// TIA Portal V21 export
// export: Created 2026-11-10T19:11:41.578579Z, ExportSetting WithDefaults, DisplayName Totally Integrated Automation Portal, DisplayVersion V21 Update 3, DisplayName STEP 7 Professional, DisplayVersion V21 Update 3, DisplayName STEP 7 Safety, DisplayVersion V21, DisplayName Tech WebApplication, DisplayVersion V21, DisplayName WinCC Basic/Comfort/Advanced, DisplayVersion V21 Update 3, DisplayName WinCC Unified, DisplayVersion V21 Update 3
DATA_BLOCK "DB_USEND_SFB"   // DB52
// stored: AutoNumber true, DBAccessibleFromOPCUA true, DBAccessibleFromWebserver true, InstanceOfName USEND_SFB, OfSystemLibElement USEND, OfSystemLibVersion 1.2
"USEND_SFB"
   // VAR_INPUT
   //    REQ : Bool;
   //    ID : CONN_PRG;
   //    R_ID : CONN_R_ID;
   // END_VAR
   // VAR_OUTPUT
   //    DONE : Bool;
   //    ERROR : Bool;
   //    STATUS : Word;
   // END_VAR
   // VAR_IN_OUT
   //    SD_1 : Variant;
   //    SD_2 : Variant;
   //    SD_3 : Variant;
   //    SD_4 : Variant;
   // END_VAR
   // VAR
   //    INDEX : Word;
   // END_VAR
BEGIN
END_DATA_BLOCK
